// TIA Portal V21 export
// export: Created 2026-08-21T20:18:51.3123552Z, ExportSetting None, DisplayName Totally Integrated Automation Portal, DisplayVersion V21, DisplayName STEP 7 Professional, DisplayVersion V21, DisplayName STEP 7 Safety, DisplayVersion V21, DisplayName Tech WebApplication, DisplayVersion V21, DisplayName WinCC Basic/Comfort/Advanced, DisplayVersion V21, DisplayName WinCC Professional, DisplayVersion V21, DisplayName WinCC Unified, DisplayVersion V21
ORGANIZATION_BLOCK "Cyclic interrupt"   // OB30, FBD, CyclicInterrupt
{ S7_Optimized_Access := 'TRUE' }
// stored: SetENOAutomatically false
   VAR_INPUT
      Initial_Call : Bool;   // Initial call of this OB
      Event_Count : Int;   // Events discarded
   END_VAR
BEGIN

REGION Network 1: Service
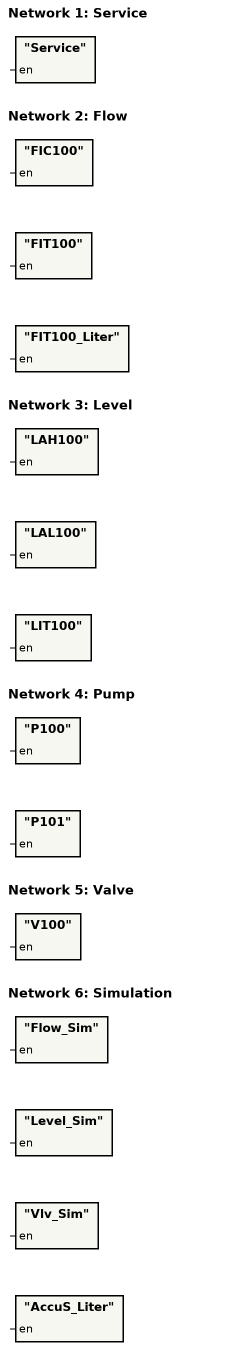
   "Service"();
END_REGION

REGION Network 2: Flow
   "FIC100"();
   "FIT100"();
   "FIT100_Liter"();
END_REGION

REGION Network 3: Level
   "LAH100"();
   "LAL100"();
   "LIT100"();
END_REGION

REGION Network 4: Pump
   "P100"();
   "P101"();
END_REGION

REGION Network 5: Valve
   "V100"();
END_REGION

REGION Network 6: Simulation
   "Flow_Sim"();
   "Level_Sim"();
   "Vlv_Sim"();
   "AccuS_Liter"();
END_REGION
END_ORGANIZATION_BLOCK
